// Restauration des valeurs rémanentes, par pages de 256 (docs/05 § 10, étape 6)
{attribute 'pack_mode' := '1'}
TYPE ST_RestoreRequest :
STRUCT
    nSeq : UDINT;
    nPage : UINT;                   // 0 = première page (efface la liste en cours)
    bLast : BOOL;                   // dernière page : appliquer
    nCount : UINT;
    aItem : ARRAY[1..256] OF ST_RetainedItem;
    sUser : STRING(24);
END_STRUCT
END_TYPE

(* stored: Version 1.1.0.1, ProductVersion 3.1.4024.12
   DUT ST_RestoreRequest: Id {5ec7c579-3382-5215-9a0f-d266cb99d2ae} *)
